Fanuc KAREL source: kd00010.KL

-- PROVISIONAL review KL for V770-1; original PC SHA256 ff8fb9ed859a4112d3b94a19d830a5047b4b390c21f79a0f876e97b761d4ae44
-- Incomplete behavior may be omitted. Consult companion uncertainty JSON. Do not deploy.
PROGRAM KD00010
%NOLOCKGROUP
VAR
  I : INTEGER
  J : INTEGER
  B : BOOLEAN
  R : REAL
  S : STRING[80]
BEGIN
  -- UNRESOLVED_PC offsets 5-12; opcodes 9D,23
  -- UNRESOLVED_PC offsets 17-21; opcodes 7F
END KD00010
